// TIA Portal project "CanvasE2E" (V19)

(* hardware
DEVICE "PLC_1"  S7-1500 station
   slot 0: "导轨_0"  Rack  6ES7 590-1***0-0AA0
   slot 1: "PLC_1"  CPU 1511-1 PN  6ES7 511-1AK01-0AB0  V2.5
      slot 3: "CPU 显示_1"  6ES7591-1AA00-0AA0
      slot 32768: "PROFINET 接口_1"  X1
         slot 32769: "端口_1"  X1 P1
         slot 32770: "端口_2"  X1 P2
*)

// ===== PLC "PLC_1"  CPU 1511-1 PN =====

TYPE "UDT_DriverState"
// AF UDT: driver runtime state
//  source_id: prj_g5_real
//  af_profile: SIEMENS_AF_BASIC_FOLDER_V19
//  template_sha256: sha256:af_basic_folder_v19_template_unbound
//  ir_sha256: sha256:f4a78f43dcfff6ab790fc68df629729a1518b66d91aee8b8684e9038a83dc351
//  deterministic semantic output: no timestamps in this file
   STRUCT
      state : Int;
      elapsed_ms : Time;
      error_id : Int;
      q_extend : Bool;
      q_retract : Bool;
   END_STRUCT;
END_TYPE

DATA_BLOCK "DB_Sequence"   // DB1
{ S7_Optimized_Access := 'TRUE' }
VERSION : 0.1
// AF instance DB for FB_Sequence (explicit, not inferred from a name)
//  source_id: prj_g5_real
//  af_profile: SIEMENS_AF_BASIC_FOLDER_V19
//  template_sha256: sha256:af_basic_folder_v19_template_unbound
//  ir_sha256: sha256:f4a78f43dcfff6ab790fc68df629729a1518b66d91aee8b8684e9038a83dc351
//  deterministic semantic output: no timestamps in this file
// stored: InstanceOfName FB_Sequence
"FB_Sequence"
BEGIN
END_DATA_BLOCK

FUNCTION_BLOCK "PumpCtrl"   // FB1, SCL
{ S7_Optimized_Access := 'TRUE' }
   VAR_INPUT
      Start : Bool;
   END_VAR
   VAR_OUTPUT
      RunOut : Bool;
   END_VAR
   VAR
      Running : Bool;
   END_VAR
BEGIN
       // Network 1: Self-holding logic
       IF #Start THEN
           #Running := TRUE;
       END_IF;
       #RunOut := #Running;
END_FUNCTION_BLOCK

FUNCTION_BLOCK "FB_Drivers"   // FB2, SCL
{ S7_Optimized_Access := 'TRUE' }
// AF FB: driver command/permission interface
//  source_id: prj_g5_real
//  af_profile: SIEMENS_AF_BASIC_FOLDER_V19
//  template_sha256: sha256:af_basic_folder_v19_template_unbound
//  ir_sha256: sha256:f4a78f43dcfff6ab790fc68df629729a1518b66d91aee8b8684e9038a83dc351
//  deterministic semantic output: no timestamps in this file
   VAR_INPUT
      CM1_CmdExtend : Bool;   // binding=None
      CM1_CmdRetract : Bool;   // binding=None
      CM1_Reset : Bool;   // binding=None
      CM1_SafetyPermit : Bool;   // binding=None
      CM1_SensorIn : Bool;   // binding=None
      CM1_SensorOut : Bool;   // binding=None
   END_VAR
   VAR_OUTPUT
      CM1_Busy : Bool;   // writer=FB_Cylinder
      CM1_Error : Bool;   // writer=FB_Cylinder
      CM1_ErrorID : Int;   // writer=FB_Cylinder
      CM1_Q_Extend : Bool;   // writer=FB_Cylinder
      CM1_Q_Retract : Bool;   // writer=FB_Cylinder
   END_VAR
BEGIN
   // Reverse outputs are interlocked by arbitrate_single_writer().
   // source_id: CM1 ; move_timeout_ms := 3000;
END_FUNCTION_BLOCK

FUNCTION_BLOCK "FB_Sequence"   // FB3, SCL
{ S7_Optimized_Access := 'TRUE' }
// AF FB: deterministic SFC-like step state machine
//  source_id: prj_g5_real
//  af_profile: SIEMENS_AF_BASIC_FOLDER_V19
//  template_sha256: sha256:af_basic_folder_v19_template_unbound
//  ir_sha256: sha256:f4a78f43dcfff6ab790fc68df629729a1518b66d91aee8b8684e9038a83dc351
//  deterministic semantic output: no timestamps in this file
   VAR_INPUT
      CmdStart : Bool;   // unbound logical signal
      HoldDone : Bool;   // unbound logical signal
      Reset : Bool;   // unbound logical signal
      SensorIn : Bool;   // unbound logical signal
      SensorOut : Bool;   // unbound logical signal
   END_VAR
   VAR
      stepCurrent : Int;
      stepElapsed_ms : Time;
      minDuration_ms : Time;
   END_VAR
BEGIN
   // Scan order: FREEZE_INPUT_SNAPSHOT -> EVALUATE_TYPED_GUARDS -> RESOLVE_PRIORITY_AND_EXCLUSIVITY -> ATOMIC_TRANSITION -> COMPOSE_ACTIONS -> ARBITRATE_SINGLE_WRITER -> TICK_DRIVER_FSMS -> EMIT_OUTPUTS_AND_ALARMS
   CASE #stepCurrent OF
       0: // source_id: S0 (IDLE)
           #minDuration_ms := T#0ms; // source_id: S0
           // guard T0: #CmdStart -> S1
           ;
       1: // source_id: S1 (EXTEND)
           #minDuration_ms := T#0ms; // source_id: S1
           // timeout_ms := 500; // source_id: S1
           // action CmdExtend := True; // source_id: S1
           // guard T1: #SensorOut -> S2
           ;
       2: // source_id: S2 (HOLD)
           #minDuration_ms := T#1000ms; // source_id: S2
           // timeout_ms := 5000; // source_id: S2
           // guard T2: #HoldDone -> S3
           ;
       3: // source_id: S3 (RETRACT)
           #minDuration_ms := T#0ms; // source_id: S3
           // timeout_ms := 500; // source_id: S3
           // action CmdRetract := True; // source_id: S3
           // guard T3: #SensorIn -> S4
           ;
       4: // source_id: S4 (DONE)
           #minDuration_ms := T#0ms; // source_id: S4
           // guard T4: NOT (#CmdStart) -> S0
           ;
       5: // source_id: FAULT (FAULT)
           #minDuration_ms := T#0ms; // source_id: FAULT
           // guard T5: #Reset -> S0
           ;
   END_CASE;
END_FUNCTION_BLOCK

ORGANIZATION_BLOCK "Main"   // OB1, LAD, ProgramCycle
TITLE = "Main Program Sweep (Cycle)"
{ S7_Optimized_Access := 'TRUE' }
VERSION : 0.1
   VAR_INPUT
      Initial_Call : Bool;   // Initial call of this OB
      Remanence : Bool;   // =True, if remanent data are available
   END_VAR
BEGIN
END_ORGANIZATION_BLOCK